FUNCTION_BLOCK FB_PID EXTENDS FB_Device
(*
	PID controller with ratio mode, for flow, level, pressure and temperature loops.
	
	Loop modes (E_PIDLoopMode), selected with ocmd/pcmd:
		Off			output = cfg.outputOff
		OpenLoop	output = manual output
		Setpoint	PID on the local setpoint
		Ratio		PID on setpoint = ratio x wildValue + cfg.ratioBias, e.g. dosing flow
					proportional to a main flow
	
	Device mode decides who sets the values: in Manual the operator (ocmd, opValues),
	in Auto the program (Off(), OpenLoop(x), Setpoint(x), Ratio(x) to change mode,
	SetOutput, SetSetpoint, SetRatio to change a value without changing mode).
	
	Bumpless: in Off and OpenLoop the integral tracks the output, and with
	cfg.setpointTracksPv the setpoint follows the PV. Anti-windup stops integrating
	while the output is limited. Derivative acts on the PV, filtered.
	If inpPvBad is TRUE in closed loop, the output is held and the loop faults.
*)
VAR_INPUT
	{attribute 'OPC.UA.DA' := '1'}
	{attribute 'OPC.UA.DA.StructuredType' := '1'}
	cfg					: ST_PIDConfiguration; //configuration
	
	{attribute 'OPC.UA.DA' := '1'}
	ocmd				: E_PIDCommand; //operator command
	{attribute 'OPC.UA.DA' := '1'}
	{attribute 'OPC.UA.DA.StructuredType' := '1'}
	opValues			: ST_PIDOperatorValues; //operator setpoint, ratio and manual output (Manual mode)
	
	(* External inputs
	----------------------------------------------------------------------------------------------------*)
	pv					: LREAL; //process value, e.g. FB_AnalogInput.sts.value
	wildValue			: LREAL; //wild (uncontrolled) value for Ratio mode, e.g. main flow
	inpPvBad			: BOOL; //PV signal is bad, e.g. NOT FB_AnalogInput.sts.valid
END_VAR
VAR_OUTPUT
	{attribute 'OPC.UA.DA' := '1'}
	{attribute 'OPC.UA.DA.Access' := '1'}
	out					: LREAL; //controller output in %, e.g. to FB_ActuatorModulating.SetPosition
	
	{attribute 'OPC.UA.DA' := '1'}
	{attribute 'OPC.UA.DA.Access' := '1'}
	{attribute 'OPC.UA.DA.StructuredType' := '1'}
	sts					: ST_PIDStatus;
	
	{attribute 'OPC.UA.DA' := '1'}
	{attribute 'OPC.UA.DA.Access' := '1'}
	{attribute 'OPC.UA.DA.StructuredType' := '1'}
	fault				: ST_PIDFault;
END_VAR
VAR
	//Command processing
	pcmd				: E_PIDCommand; //program command
	pcmdLast			: E_PIDCommand;
	ocmdLast			: E_PIDCommand;
	cmdReceived			: E_PIDCommand; //command accepted this scan
	pSetpoint			: LREAL; //program setpoint
	pRatio				: LREAL; //program ratio
	pOutput				: LREAL; //program manual output
	
	//Controller state
	integral			: LREAL; //integral term in % output
	pvLast				: LREAL; //PV on the previous scan, for the derivative
	pvSlopeFiltered		: LREAL; //filtered dPV/stepTime
	firstScan			: BOOL := TRUE; //no derivative on the first scan
	
	//Alarms
	deviationAlarm		: FB_LimitAlarm; //|error| above deviationLimit
	
	//Timers
	deltaTime			: FB_DeltaTime; //scan time for the controller
	
	resetFault			: BOOL;
END_VAR
VAR CONSTANT
	LIMIT_BAND			: LREAL := 1E-6; //output within this of a limit counts as at the limit (floating point rounding)
END_VAR

SUPER^();

Device();
ProcessInputs();
ProcessCommands();
StateMachine();
HandleFaults();
ControlOutputs();
StatusOut();

METHOD PROTECTED ControlOutputs //PID calculation and output limits
VAR
	direction	: LREAL; //+1 reverse acting, -1 direct acting
	target		: LREAL; //output before the rate limit
	pvSlope		: LREAL; //unfiltered dPV/stepTime
	tiSec		: LREAL; //integral time in s
	tdSec		: LREAL; //derivative time in s
	tfSec		: LREAL; //derivative filter in s
	stepTime			: LREAL; //scan time in s
END_VAR
stepTime		:= deltaTime.seconds;
tiSec	:= TIME_TO_LREAL(cfg.ti) / 1000.0;
tdSec	:= TIME_TO_LREAL(cfg.td) / 1000.0;
tfSec	:= TIME_TO_LREAL(cfg.tdFilter) / 1000.0;
direction := SEL(cfg.directActing, 1.0, -1.0);

//Derivative on the PV (not the error) so setpoint changes don't kick the output
IF firstScan OR stepTime <= 0 THEN
	pvSlope := 0;
	firstScan := FALSE;
ELSE
	pvSlope := (sts.pv - pvLast) / stepTime;
END_IF
pvLast := sts.pv;
IF tfSec > 0 THEN
	pvSlopeFiltered := pvSlopeFiltered + stepTime / (tfSec + stepTime) * (pvSlope - pvSlopeFiltered);
ELSE
	pvSlopeFiltered := pvSlope;
END_IF

sts.pTerm := direction * cfg.kp * sts.error;
sts.dTerm := -direction * cfg.kp * tdSec * pvSlopeFiltered;

CASE sts.loopMode OF
	
	E_PIDLoopMode.Setpoint, E_PIDLoopMode.Ratio:
		//Anti-windup: only integrate when it moves the output away from a limit it is not at
		IF tiSec > 0 AND NOT ((sts.output >= cfg.outputMax - LIMIT_BAND AND direction * sts.error > 0)
							 OR (sts.output <= cfg.outputMin + LIMIT_BAND AND direction * sts.error < 0)) THEN
			integral := integral + direction * cfg.kp * sts.error * stepTime / tiSec;
		END_IF
		IF tiSec <= 0 THEN
			integral := 0;
		END_IF
		integral := LIMIT(cfg.outputMin - sts.pTerm - sts.dTerm, integral, cfg.outputMax - sts.pTerm - sts.dTerm);
		target := sts.pTerm + integral + sts.dTerm;
		
	E_PIDLoopMode.OpenLoop:
		target := sts.manualOutput;
		
ELSE // Off
	target := cfg.outputOff;
	
END_CASE

target := LIMIT(cfg.outputMin, target, cfg.outputMax);
//Snap to the limit so it is exact after rounding
IF target >= cfg.outputMax - LIMIT_BAND THEN
	target := cfg.outputMax;
ELSIF target <= cfg.outputMin + LIMIT_BAND THEN
	target := cfg.outputMin;
END_IF
IF sts.loopMode = E_PIDLoopMode.Off THEN
	target := cfg.outputOff; // outputOff may be outside the control range
END_IF

//Rate limit
IF cfg.outputRateLimit > 0 AND sts.closedLoop THEN
	sts.output := sts.output + LIMIT(-cfg.outputRateLimit * stepTime, target - sts.output, cfg.outputRateLimit * stepTime);
ELSE
	sts.output := target;
END_IF

//Bumpless transfer: outside closed loop the integral tracks the output
IF NOT sts.closedLoop THEN
	integral := sts.output - sts.pTerm - sts.dTerm;
	IF sts.loopMode = E_PIDLoopMode.OpenLoop THEN
		pOutput := opValues.output := sts.manualOutput;
	END_IF
ELSE
	//Manual output follows the loop so switching to OpenLoop does not bump
	pOutput := opValues.output := sts.manualOutput := sts.output;
END_IF
sts.iTerm := integral;
END_METHOD

METHOD PROTECTED Device //map cfg to FB_Device and FB_Device to sts
// to FB device
opTimeout  			 := cfg.opTimeout;
opTimeoutEnable 	 := cfg.opTimeoutEnable;
opActivity 			 := ocmd <> E_PIDCommand.None;

// from FB device
sts.mode	   		 := mode;
sts.modeAuto   		 := sts.mode = E_SystemMode.Auto;
sts.modeManual 		 := sts.mode = E_SystemMode.Manual;
sts.manualOvrde		 := ctrl.manualOvrde;
sts.bypass 	   		 := ctrl.bypass;
sts.sim		   		 := ctrl.sim;
sts.parentConfigured := parentConfigured;
END_METHOD

METHOD PROTECTED HandleFaults
fault.pvBad S= inpPvBad AND sts.closedLoop;
//fault.ocmdNOK; // Set in ProcessCommands
//fault.pcmdNOK; // Set in ProcessCommands

(* ----- Handle Reset ----- *)
IF resetFault THEN
	fault.ocmdNOK R= TRUE;
	fault.pcmdNOK R= TRUE;
	fault.pvBad R= NOT inpPvBad; // only clears once the PV is good again
END_IF
resetFault := FALSE;

(* ----- Map Fault Id ----- *)
fault.id.0 := fault.ocmdNOK;
fault.id.1 := fault.pcmdNOK;
fault.id.2 := fault.pvBad;

(* ----- Map Fault Text ----- *)
IF fault.ocmdNOK THEN		fault.text := 'Operator command in Auto is not allowed';
ELSIF fault.pcmdNOK THEN	fault.text := 'Program command in Manual is not allowed';
ELSIF fault.pvBad THEN		fault.text := CONCAT(cfg.loopId, ' PV bad, output held');
ELSE fault.text := '';
END_IF

(* ----- Set Active ----- *)
fault.active := fault.id > 0;
END_METHOD

METHOD PUBLIC Off //loop off, output to cfg.outputOff
pcmd := E_PIDCommand.Off;
END_METHOD

METHOD PROTECTED ProcessCommands
//Check for new valid commands
IF ctrl.reset THEN
	PrvReset();
ELSIF ocmd <> E_PIDCommand.None THEN
	IF sts.modeManual THEN
		cmdReceived := ocmd;
	ELSE
		fault.ocmdNOK := TRUE;
	END_IF
ELSIF pcmd <> E_PIDCommand.None THEN
	IF sts.modeAuto THEN
		cmdReceived := pcmd;
	ELSE
		fault.pcmdNOK := TRUE;
	END_IF
END_IF

//Values: the operator owns them in Manual, the program in Auto. The other side is
//kept equal, so switching mode does not change anything.
IF sts.modeManual THEN
	pSetpoint			:= opValues.setpoint;
	pRatio				:= opValues.ratio;
	pOutput				:= opValues.output;
ELSE
	opValues.setpoint	:= pSetpoint;
	opValues.ratio		:= pRatio;
	opValues.output		:= pOutput;
END_IF
sts.localSetpoint	:= pSetpoint;
sts.ratio			:= pRatio;
sts.manualOutput	:= pOutput;
sts.localSetpoint	:= LIMIT(cfg.setpointMin, sts.localSetpoint, cfg.setpointMax);
sts.ratio			:= LIMIT(cfg.ratioMin, sts.ratio, cfg.ratioMax);
sts.manualOutput	:= LIMIT(cfg.outputMin, sts.manualOutput, cfg.outputMax);

CASE cmdReceived OF
	E_PIDCommand.Off:
		PrvOff();
	E_PIDCommand.OpenLoop:
		PrvOpenLoop();
	E_PIDCommand.Setpoint:
		PrvSetpoint();
	E_PIDCommand.Ratio:
		PrvRatio();
END_CASE

//Save last commands
IF pcmd <> E_PIDCommand.None THEN
	pcmdLast := pcmd;
END_IF
IF ocmd <> E_PIDCommand.None THEN
	ocmdLast := ocmd;
END_IF

//Clear commands every scan
cmdReceived	:= E_PIDCommand.None;
pcmd		:= E_PIDCommand.None;
ocmd		:= E_PIDCommand.None;
ctrl.reset	:= FALSE;
END_METHOD

METHOD PROTECTED ProcessInputs
deltaTime();

sts.pv			:= pv;
sts.wildValue	:= wildValue;
END_METHOD

METHOD PROTECTED PrvReset //Reset the loop
resetFault S= TRUE;
END_METHOD

METHOD PUBLIC SetOutput //program: change the manual output without changing mode
VAR_INPUT
	output		: LREAL; //output in %
END_VAR
pOutput := output;
END_METHOD

METHOD PUBLIC SetRatio //program: change the ratio without changing mode
VAR_INPUT
	ratio		: LREAL; //ratio
END_VAR
pRatio := ratio;
END_METHOD

METHOD PUBLIC SetSetpoint //program: change the setpoint without changing mode
VAR_INPUT
	setpoint	: LREAL; //setpoint in PV units
END_VAR
pSetpoint := setpoint;
END_METHOD

METHOD PROTECTED StateMachine //active setpoint and error
//A bad PV in closed loop holds the current output in OpenLoop
IF inpPvBad AND sts.closedLoop THEN
	fault.pvBad S= TRUE;
	pOutput := opValues.output := sts.output;
	sts.manualOutput := sts.output;
	sts.loopMode := E_PIDLoopMode.OpenLoop;
END_IF

sts.closedLoop := sts.loopMode = E_PIDLoopMode.Setpoint OR sts.loopMode = E_PIDLoopMode.Ratio;

CASE sts.loopMode OF
	E_PIDLoopMode.Ratio:
		sts.setpoint := LIMIT(cfg.setpointMin, sts.ratio * sts.wildValue + cfg.ratioBias, cfg.setpointMax);
	E_PIDLoopMode.Setpoint:
		sts.setpoint := sts.localSetpoint;
ELSE
	//Open loop: setpoint follows the PV so closing the loop does not bump
	IF cfg.setpointTracksPv THEN
		pSetpoint := opValues.setpoint := sts.localSetpoint := LIMIT(cfg.setpointMin, sts.pv, cfg.setpointMax);
	END_IF
	sts.setpoint := sts.localSetpoint;
END_CASE

sts.error := sts.setpoint - sts.pv;

deviationAlarm(value := ABS(sts.error), threshold := cfg.deviationLimit, highAlarm := TRUE,
			   enable := cfg.deviationEnable AND sts.closedLoop, deadband := cfg.deviationLimit * 0.1,
			   delay := cfg.deviationDelay, latch := FALSE, reset := FALSE);
END_METHOD

METHOD PROTECTED StatusOut //Set output status information
sts.saturatedHigh	:= sts.closedLoop AND sts.output >= cfg.outputMax;
sts.saturatedLow	:= sts.closedLoop AND sts.output <= cfg.outputMin;
sts.deviationAlarm	:= deviationAlarm.active;
out					:= sts.output;
END_METHOD

METHOD PUBLIC Setpoint //closed loop on a setpoint
VAR_INPUT
	value		: LREAL; //setpoint in PV units
END_VAR
pSetpoint := value;
pcmd := E_PIDCommand.Setpoint;
END_METHOD

METHOD PUBLIC Ratio //closed loop on ratio x wildValue + cfg.ratioBias
VAR_INPUT
	value		: LREAL; //ratio
END_VAR
pRatio := value;
pcmd := E_PIDCommand.Ratio;
END_METHOD

METHOD PUBLIC OpenLoop //open loop at a fixed output
VAR_INPUT
	value		: LREAL; //output in %
END_VAR
pOutput := value;
pcmd := E_PIDCommand.OpenLoop;
END_METHOD

METHOD PROTECTED PrvOff
sts.loopMode := E_PIDLoopMode.Off;
END_METHOD

METHOD PROTECTED PrvOpenLoop
sts.loopMode := E_PIDLoopMode.OpenLoop;
END_METHOD

METHOD PROTECTED PrvSetpoint
IF inpPvBad THEN // cannot close the loop on a bad PV
	fault.pvBad S= TRUE;
ELSE
	sts.loopMode := E_PIDLoopMode.Setpoint;
END_IF
END_METHOD

METHOD PROTECTED PrvRatio
IF inpPvBad THEN // cannot close the loop on a bad PV
	fault.pvBad S= TRUE;
ELSE
	sts.loopMode := E_PIDLoopMode.Ratio;
END_IF
END_METHOD

END_FUNCTION_BLOCK

(* stored: Version 1.1.0.1, ProductVersion 3.1.4024.12
   POU FB_PID: Id {c0565bc6-ce91-4676-8689-a6a4bae45924}, SpecialFunc None
   Folder Protected: Id {df9d7a5f-dca8-4f53-91b0-517d713c4c5e}
   Folder Commands: Id {8fcef680-1800-4baf-a415-bf012222821a}
   Folder Logic: Id {c3db8777-1fb3-47e6-8373-d722144aa706}
   Folder Public: Id {a660de5a-cdd3-4117-aa5a-d90de0461f5e}
   Folder Commands: Id {437152d1-5f8b-4d80-be40-f40f5c8cd146}
   Folder Control: Id {9db9fc39-7e11-444b-9b33-660d86c53f99}
   Method ControlOutputs: Id {568b6f2e-991b-4036-98bf-610feb1f91b8}
   Method Device: Id {359421ee-ae5d-4589-b7e0-abe53108efba}
   Method HandleFaults: Id {35e9c03b-52e6-4791-9977-6a2b6cdcffe3}
   Method Off: Id {a15d9aad-794b-4db9-a2eb-520c09d45ef3}
   Method ProcessCommands: Id {16672a96-a407-4e2c-be5b-1023dfd456c0}
   Method ProcessInputs: Id {a9dcf913-7ac9-4d5d-be38-92cd3150115f}
   Method PrvReset: Id {56dc3802-ad3e-49f7-bf88-68657f64f0b5}
   Method SetOutput: Id {030395d2-e421-4926-9461-a1ab9df16968}
   Method SetRatio: Id {6fc2908a-ff22-4554-9d89-61e40629c84a}
   Method SetSetpoint: Id {17329377-891f-47d0-a901-d0537959adf6}
   Method StateMachine: Id {a3e7e3c1-3042-40c4-8ab9-adee7a2fbecc}
   Method StatusOut: Id {757cfed1-89b5-4407-8ffe-70f651f49e19}
   Method Setpoint: Id {752fe3e6-8416-4b02-89de-3fd761e7e2e3}
   Method Ratio: Id {1b5cc355-df22-4c92-89be-33f7d5aa0123}
   Method OpenLoop: Id {904d7c5f-542d-4d58-8c0f-1a78aa230b43}
   Method PrvOff: Id {f11db683-15d0-4b32-80e6-4c8d8c965ac0}
   Method PrvOpenLoop: Id {48935ea2-7e3a-47a1-848d-9d52816a41fb}
   Method PrvSetpoint: Id {4f30a4fc-dcb7-4080-9ce3-349dcf2b3a27}
   Method PrvRatio: Id {a7dfa6a3-f805-49b6-a383-12f7ba9788aa} *)
